FUNCTION_BLOCK GATE_CYCLE
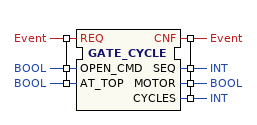
  EVENT_INPUT
    REQ WITH OPEN_CMD, AT_TOP;
  END_EVENT
  EVENT_OUTPUT
    CNF WITH SEQ, MOTOR, CYCLES;
  END_EVENT
  VAR_INPUT
    OPEN_CMD : BOOL;
    AT_TOP : BOOL;
  END_VAR
  VAR_OUTPUT
    SEQ : INT;
    MOTOR : BOOL;
    CYCLES : INT;
  END_VAR
  VAR
    K : INT;
  END_VAR
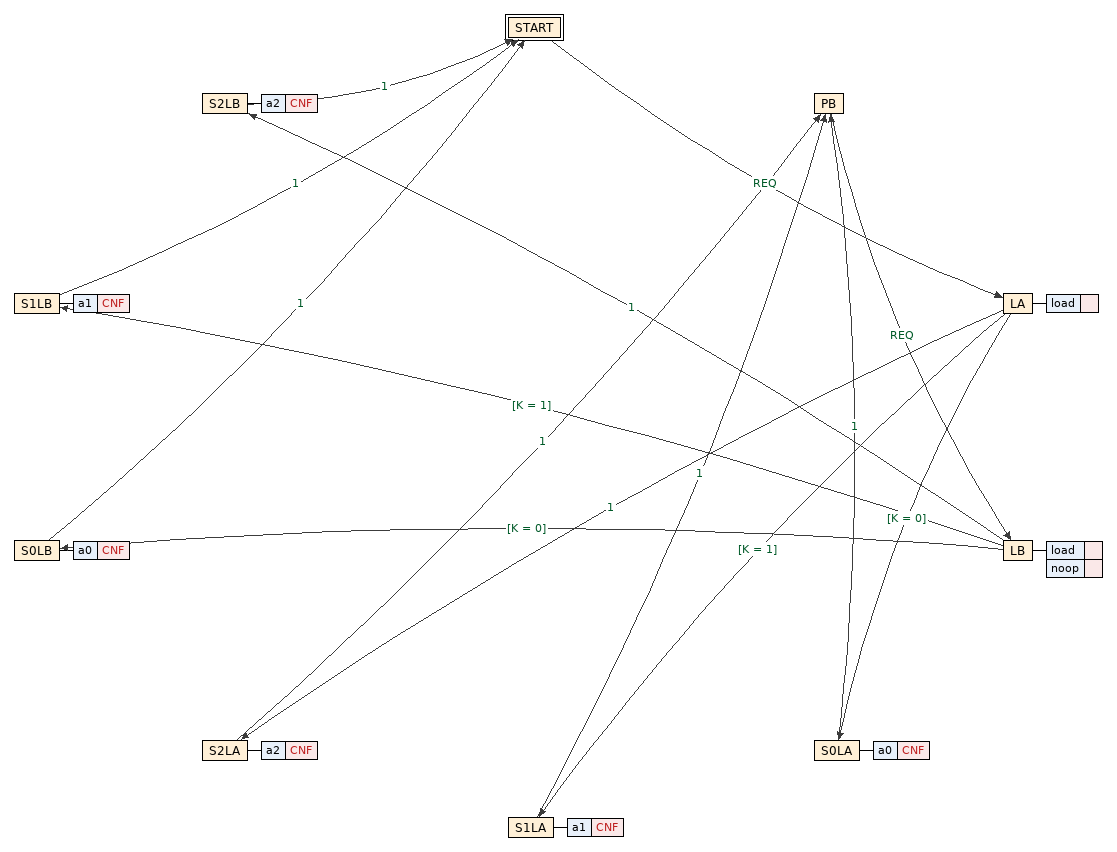
  EC_STATES
    START;
    PB;
    LA : load;
    LB : load, noop;
    S0LA : a0 -> CNF;
    S1LA : a1 -> CNF;
    S2LA : a2 -> CNF;
    S0LB : a0 -> CNF;
    S1LB : a1 -> CNF;
    S2LB : a2 -> CNF;
  END_STATES
  EC_TRANSITIONS
    START TO LA := REQ;
    PB TO LB := REQ;
    LA TO S0LA := [K = 0];
    S0LA TO PB := 1;
    LA TO S1LA := [K = 1];
    S1LA TO PB := 1;
    LA TO S2LA := 1;
    S2LA TO PB := 1;
    LB TO S0LB := [K = 0];
    S0LB TO START := 1;
    LB TO S1LB := [K = 1];
    S1LB TO START := 1;
    LB TO S2LB := 1;
    S2LB TO START := 1;
  END_TRANSITIONS
  ALGORITHM load IN ST:
K := SEQ;
  END_ALGORITHM
  ALGORITHM noop IN ST:
CYCLES := CYCLES;
  END_ALGORITHM
  ALGORITHM a0 IN ST:
MOTOR := FALSE;
IF OPEN_CMD THEN SEQ := 1; END_IF;
  END_ALGORITHM
  ALGORITHM a1 IN ST:
MOTOR := TRUE;
IF AT_TOP THEN SEQ := 2; END_IF;
  END_ALGORITHM
  ALGORITHM a2 IN ST:
MOTOR := FALSE;
CYCLES := CYCLES + 1;
SEQ := 0;
  END_ALGORITHM
END_FUNCTION_BLOCK
